(* IEC 61131-3 sources: tia-guard/examples/twincat3-generation/motor/sources, 5 files *)

(* ---- ST_MotorStatus.declaration.st ---- *)
TYPE ST_MotorStatus :
STRUCT
    Running : BOOL;
    Faulted : BOOL;
    CycleCount : UDINT;
END_STRUCT
END_TYPE

(* ---- GVL_Signals.declaration.st ---- *)
VAR_GLOBAL
    Start : BOOL;
    Stop : BOOL;
    Fault : BOOL;
    Reset : BOOL;
    Status : ST_MotorStatus;
END_VAR

(* ---- FB_Motor.declaration.st ---- *)
FUNCTION_BLOCK FB_Motor
VAR_INPUT
    Start : BOOL;
    Stop : BOOL;
    Fault : BOOL;
    Reset : BOOL;
END_VAR
VAR_OUTPUT
    Status : ST_MotorStatus;
END_VAR

(* ---- FB_Motor.implementation.st ---- *)
Status.CycleCount := Status.CycleCount + 1;
IF Fault THEN
    Status.Faulted := TRUE;
ELSIF Reset THEN
    Status.Faulted := FALSE;
END_IF;
IF Stop OR Status.Faulted THEN
    Status.Running := FALSE;
ELSIF Start THEN
    Status.Running := TRUE;
END_IF;

(* ---- MAIN.declaration.st ---- *)
PROGRAM MAIN
VAR
    Motor : FB_Motor;
END_VAR
